(*
SPDX-FileCopyrightText: © 2026 Oleksandr Tiutyk <trofimich@gmail.com>
SPDX-License-Identifier: MIT
License: https://opensource.org/license/mit
*)
(*!
<summary>Owns one captured logger call independently of caller buffers.</summary>
*)
TYPE LOGGER_CAPTURED_MESSAGE :
STRUCT
	Category : TOF_Core.LOG_CATEGORY;
	Message : TOF_Core.ERROR_MESSAGE;
	HasMessageNumber : BOOL;
	MessageNumber : ULINT;
END_STRUCT
END_TYPE

(* stored: Version 1.1.0.1
   DUT LOGGER_CAPTURED_MESSAGE: Id {d18ab71e-0a07-4199-887c-920fd6ce0777} *)
